// TIA Portal V20 export
Screen "200FX1Layout"  1276x673
  ScreenItem "Line_Header_X0_Y64" at 0,64 size 1276x0  Type=HmiLine
  ScreenItem "permanentareaborderrectangle" at 0,0 size 0x0  Type=HmiRectangle
  ScreenItem "Button_Back" at 2,2 size 90x60  Type=HmiButton
  ScreenItem "Move_Legend" at 1182,2 size 90x60  Type=HmiButton
  ScreenItem "Fusszeile_Button_ManualOPMode1_2" at 279,2 size 90x60  Type=HmiButton
  ScreenItem "文本域_3" at 1107,71 size 139x22  Type=HmiTextBox
  ScreenItem "LSicar_Valve8Pos_LeftHomeRightWork_WithPB_5" at 1099,95 size 160x53  Type=HmiFaceplateContainer
  ScreenItem "文本域_1" at 1107,160 size 156x23  Type=HmiTextBox
  ScreenItem "LSicar_Valve8Pos_LeftHomeRightWork_WithPB_1" at 1099,183 size 160x53  Type=HmiFaceplateContainer
  ScreenItem "文本域_2" at 1107,246 size 135x23  Type=HmiTextBox
  ScreenItem "LSicar_Valve8Pos_LeftHomeRightWork_WithPB_2" at 1099,271 size 160x53  Type=HmiFaceplateContainer
  ScreenItem "文本域_22" at 1124,475 size 104x23  Type=HmiTextBox
  ScreenItem "面板容器_23" at 1171,508 size 96x32  Type=HmiFaceplateContainer
  ScreenItem "面板容器_22" at 1061,508 size 96x32  Type=HmiFaceplateContainer
  ScreenItem "面板容器_2" at 1090,4 size 88x58  Type=HmiFaceplateContainer
  ScreenItem "OPMode1_Blocked" at 1164,6 size 14x14  Type=HmiGraphicView
  ScreenItem "OPMode4_Foreground_Blocked" at 982,13 size 88x58  Type=HmiGraphicView
  ScreenItem "Fusszeile_Button_ManualOPMode1_1" at 95,2 size 90x60  Type=HmiButton
  ScreenItem "LSicar_Valve8Pos_LeftHomeRightWork_WithPB_4" at 1099,356 size 160x53  Type=HmiFaceplateContainer
  ScreenItem "文本域_4" at 1107,330 size 139x22  Type=HmiTextBox
  ScreenItem "Button_Back_1" at 1180,606 size 90x60  Type=HmiButton
  ScreenItem "面板容器_1" at 424,537 size 62x46  Type=HmiFaceplateContainer
  ScreenItem "面板容器_3" at 951,383 size 59x50  Type=HmiFaceplateContainer
  ScreenItem "Faceplate container_1" at 296,523 size 69x45  Type=HmiFaceplateContainer
  ScreenItem "面板容器_9" at 684,588 size 172x60  Type=HmiFaceplateContainer
  ScreenItem "面板容器_14" at 33,195 size 58x51  Type=HmiFaceplateContainer
  ScreenItem "Faceplate container_3" at 678,183 size 59x48  Type=HmiFaceplateContainer
  ScreenItem "Faceplate container_4" at 439,192 size 59x47  Type=HmiFaceplateContainer
  ScreenItem "面板容器_20" at 534,612 size 150x51  Type=HmiFaceplateContainer
  ScreenItem "Graphic view_1" at 20,214 size 860x259  Type=HmiGraphicView
  ScreenItem "Line_9" at 559,146 size 94x182  Type=HmiLine
  ScreenItem "面板容器_10" at 498,116 size 153x58  Type=HmiFaceplateContainer
  ScreenItem "Line_2" at 703,221 size 20x91  Type=HmiLine
  ScreenItem "Line_5" at 753,170 size 92x151  Type=HmiLine
  ScreenItem "Line_3" at 514,184 size 62x132  Type=HmiLine
  ScreenItem "Line_17" at 109,190 size 171x117  Type=HmiLine
  ScreenItem "Line_6" at 752,357 size 177x7  Type=HmiLine
  ScreenItem "Line_10" at 558,396 size 165x104  Type=HmiLine
  ScreenItem "Line_13" at 603,398 size 127x171  Type=HmiLine
  ScreenItem "Line_1" at 445,359 size 219x135  Type=HmiLine
  ScreenItem "Line_8" at 328,395 size 248x99  Type=HmiLine
  ScreenItem "Line_18" at 218,401 size 62x96  Type=HmiLine
  ScreenItem "Line_16" at 71,325 size 85x136  Type=HmiLine
  ScreenItem "面板容器_6" at 914,208 size 149x54  Type=HmiFaceplateContainer
  ScreenItem "面板容器_5" at 12,502 size 143x50  Type=HmiFaceplateContainer
  ScreenItem "面板容器_4" at 520,522 size 62x46  Type=HmiFaceplateContainer
  ScreenItem "Faceplate container_2" at 188,522 size 60x47  Type=HmiFaceplateContainer
  ScreenItem "Fusszeile_Button_ManualOPMode1_3" at 187,2 size 90x60  Type=HmiButton
  ScreenItem "Fusszeile_Button_ManualOPMode1_4" at 997,2 size 90x60  Type=HmiButton
  ScreenItem "Fusszeile_Button_ManualOPMode1_5" at 902,1 size 90x60  Type=HmiButton
  ScreenItem "文本域_19" at 168,499 size 100x20  Type=HmiTextBox
  ScreenItem "文本域_6" at 12,461 size 140x40  Type=HmiTextBox
  ScreenItem "文本域_7" at 277,500 size 100x20  Type=HmiTextBox
  ScreenItem "文本域_8" at 398,494 size 100x40  Type=HmiTextBox
  ScreenItem "文本域_9" at 513,501 size 100x20  Type=HmiTextBox
  ScreenItem "文本域_10" at 534,571 size 140x40  Type=HmiTextBox
  ScreenItem "文本域_11" at 684,565 size 140x20  Type=HmiTextBox
  ScreenItem "文本域_12" at 931,343 size 100x40  Type=HmiTextBox
  ScreenItem "文本域_13" at 503,94 size 140x20  Type=HmiTextBox
  ScreenItem "文本域_14" at 936,-172 size 140x40  Type=HmiTextBox
  ScreenItem "文本域_15" at 914,166 size 140x40  Type=HmiTextBox
  ScreenItem "文本域_16" at 12,175 size 100x20  Type=HmiTextBox
  ScreenItem "文本域_17" at 415,169 size 100x20  Type=HmiTextBox
  ScreenItem "文本域_18" at 653,160 size 100x20  Type=HmiTextBox
  ScreenItem "文本域_5" at -1,82 size 120x40  Type=HmiTextBox
  ScreenItem "Title_ScreenOverview_X390_Y2_1" at 384,5 size 510x57  Type=HmiTextBox
  ScreenItem "文本域_20" at 767,114 size 140x20  Type=HmiTextBox
  ScreenItem "面板容器_7" at 776,136 size 148x58  Type=HmiFaceplateContainer
  ScreenItem "面板容器_8" at 129,123 size 144x51  Type=HmiFaceplateContainer
  ScreenItem "文本域_21" at 129,82 size 140x40  Type=HmiTextBox
  ScreenItem "文本域_23" at 282,82 size 140x40  Type=HmiTextBox
  ScreenItem "Line_11" at 355,151 size 68x134  Type=HmiLine
  ScreenItem "Line_4" at 198,146 size 221x158  Type=HmiLine
  ScreenItem "Line_12" at 778,194 size 133x129  Type=HmiLine
  ScreenItem "文本域_24" at 913,264 size 140x20  Type=HmiTextBox
  ScreenItem "面板容器_12" at 922,286 size 148x58  Type=HmiFaceplateContainer
  ScreenItem "文本域_25" at 921,433 size 140x20  Type=HmiTextBox
  ScreenItem "面板容器_13" at 930,455 size 148x58  Type=HmiFaceplateContainer
  ScreenItem "文本域_26" at 911,548 size 140x40  Type=HmiTextBox
  ScreenItem "面板容器_15" at 914,590 size 149x54  Type=HmiFaceplateContainer
  ScreenItem "Line_14" at 754,274 size 161x75  Type=HmiLine
  ScreenItem "Line_15" at 754,367 size 166x74  Type=HmiLine
  ScreenItem "Line_7" at 746,389 size 3x173  Type=HmiLine
  ScreenItem "Line_19" at 778,386 size 132x186  Type=HmiLine
  ScreenItem "文本域_27" at -1,126 size 120x40  Type=HmiTextBox
  ScreenItem "面板容器_11" at 282,123 size 150x51  Type=HmiFaceplateContainer
  ScreenItem "Button_Back_3" at 122,606 size 90x60  Type=HmiButton
  ScreenItem "Button_Back_2" at 8,606 size 90x60  Type=HmiButton
  ScreenItem "OPMode4_Foreground_Blocked_1" at 1090,7 size 88x58  Type=HmiGraphicView
